{attribute 'qualified_only'}
{attribute 'strict'}
{attribute 'to_string'}
TYPE eShutterCommandType :
(
    NONE,           // No command
    OPEN,           // Open command (move to 100%)
    CLOSE,          // Close command (move to 0%)
	STEP_OPEN,		// Open by step 10%
	STEP_CLOSE,		// Close by step 10%
    STOP,           // Stop command
    MOVE_TO_POSITION // Move to specific position
);
END_TYPE

(* stored: Version 1.1.0.1
   DUT eShutterCommandType: Id {23be3c58-230f-4a45-8a04-cf15dcfe10a1} *)
